Staubli VAL3: mainCycle.pgx

public program mainCycle()
  local bool l_bOut
  local string l_sStr
  local num l_nVal
begin
  l_bOut=false
  do
    //*************************************************************************************************
    //Refresh the widgets of the <Page_Container_Main>：
    //*************************************************************************************************
    call db:refreshLanguage()
    call db:refreshCheckBox(db:utImg_CheckBox_a)
    call db:refreshCheckBox(db:utImg_CheckBox_b)
    call db:refreshJogMode()
    call db:refreshInfo()
    call db:refreshQuit(l_bOut)
    //
    call refreshBtn0_CaliTcp()
    //
    call refreshBtn1_AdjXY()
    //
    call refreshBtn2_Test()
    //

  until l_bOut
end
